// TwinCAT 3 PLC project MyLibrary
// Title: MyLibrary
// Company: FabioBolognesi
// Author: Fabio Bolognesi
// ProjectVersion: 0.0.0.0
// ProgramVersion: 3.1.4023.0
// libraries:
//   Tc2_Standard, * (Beckhoff Automation GmbH)
//   Tc2_System, * (Beckhoff Automation GmbH)
//   Tc2_Utilities, * (Beckhoff Automation GmbH)
//   Tc3_Module, * (Beckhoff Automation GmbH)
// project tree:
//   FUNCTION_BLOCKs/ FB_stringBuilder.TcPOU, FB_sweep.TcPOU, FB_timer.TcPOU
//   FUNCTIONs/ F_atan2.TcPOU, F_interpolateReal.TcPOU, F_interpolateTime.TcPOU, F_saturation.TcPOU, F_time2seconds.TcPOU, F_seconds2time.TcPOU
//   GLOBAL_VARIABLEs/ CONSTANTS.TcGVL, CONVERSIONS.TcGVL, PARAMETERs.TcGVL
//   STRUCTUREs/ ST_TypeSizes.TcDUT
// real-time tasks:
//   TASK PlcTask: cycle T#10ms, priority 20, ADS port 350

// ---- STRUCTUREs/ST_TypeSizes.TcDUT
TYPE ST_TypeSizes :
STRUCT
	// MEMORIA
	uiBIT		:	UINT	:=	SIZEOF(BIT);
	uiByte		:	UINT	:=	SIZEOF(BYTE);
	uiWord		:	UINT	:=	SIZEOF(WORD);
	uiDWord		:	UINT	:=	SIZEOF(DWORD);
	uiLWord		:	UINT	:=	SIZEOF(LWORD);
	
	// BOOL
	uiBool		:	UINT	:=	SIZEOF(BOOL);
	
	// UINTERI
	uiSUINT		:	UINT	:=	SIZEOF(SINT);
	uiUSUINT	:	UINT	:=	SIZEOF(USINT);
	uiUINT		:	UINT	:=	SIZEOF(UINT);
	uiUUINT		:	UINT	:=	SIZEOF(UINT);
	uiDUINT		:	UINT	:=	SIZEOF(DINT);
	uiUDUINT	:	UINT	:=	SIZEOF(UDINT);
	uiLUINT		:	UINT	:=	SIZEOF(LINT);
	uiULUINT	:	UINT	:=	SIZEOF(ULINT);
	
	// REALI
	uiReal		:	UINT	:=	SIZEOF(REAL);
	uiLReal		:	UINT	:=	SIZEOF(LREAL);
	
	// STRINGE
	
	// TEMPI E DATE
	uiTime		:	UINT	:=	SIZEOF(TIME);
	uiLTime		:	UINT	:=	SIZEOF(LTIME);
	uiDate		:	UINT	:=	SIZEOF(DATE);
	
	// MIE FUNCTION BLOCKS
	uiStringBuilder	:	UINT	:=	SIZEOF(FB_stringBuilder);
	uiTimer			:	UINT	:=	SIZEOF(FB_timer);
	
END_STRUCT
END_TYPE

// ---- GLOBAL_VARIABLEs/CONSTANTS.TcGVL
{attribute 'qualified_only'}
VAR_GLOBAL CONSTANT
	// ACCELERAZIONE DI GRAVITà
	G	:	REAL	:=	9.80665;
	
	// PI GRECO
	PI	:	REAL	:=	3.141592;
	
END_VAR

// ---- GLOBAL_VARIABLEs/CONVERSIONS.TcGVL
{attribute 'qualified_only'}
VAR_GLOBAL CONSTANT
	rTime2Seconds	:	REAL	:=	0.001;
	rSeconds2Time	:	REAL	:=	1000;
END_VAR

// ---- GLOBAL_VARIABLEs/PARAMETERs.TcGVL
{attribute 'global_init_slot' := '40001'}
{attribute 'qualified_only'}
VAR_GLOBAL CONSTANT
	// CARATTERI MASSIMI PER STRINGHE
	uiMaxCharacters	:	UINT	:=	5000;
END_VAR

// ---- FUNCTION_BLOCKs/FB_stringBuilder.TcPOU
FUNCTION_BLOCK FB_stringBuilder
VAR_INPUT
END_VAR
VAR
	bBuffer				:	ARRAY[0..PARAMETERS.uiMaxCharacters - 1] OF BYTE;
	bBufferOld			:	ARRAY[0..PARAMETERS.uiMaxCharacters - 1] OF BYTE;
	udiIndex			:	UDINT;
	udiIndexOld			:	UDINT;
	pbBuffer			:	POINTER TO BYTE		:=	ADR(bBuffer);
	pbBufferOld			:	POINTER TO BYTE		:=	ADR(bBufferOld);
END_VAR

METHOD AddChar : BOOL
VAR_INPUT
	byChar	:	BYTE;
END_VAR
IF CheckLength() THEN
	bBuffer[udiIndex]	:=	byChar;
	AddChar			:=	TRUE;
	IncrementIndex();
END_IF
END_METHOD

ACTION AddCloseBracket:
AddChar(41);
END_ACTION

ACTION AddColon:
AddChar(58);
END_ACTION

ACTION AddComma:
AddChar(44);
END_ACTION

ACTION AddDollar:
AddChar(36);
END_ACTION

ACTION AddDot:
AddChar(46);
END_ACTION

ACTION AddDoubleQuote:
AddChar(34);
END_ACTION

METHOD AddKeyValue : BOOL
VAR_INPUT
	psKey	:	POINTER TO STRING;
	psValue	:	POINTER TO STRING;
END_VAR
AddString(psKey);
AddColon();
AddString(psValue);
AddComma();
END_METHOD

ACTION AddNewLine:
AddChar(10);
END_ACTION

ACTION AddNullChar:
IF NOT CheckLength() THEN
	udiIndex	:=	PARAMETERS.uiMaxCharacters - 1;
END_IF
AddChar(0);
END_ACTION

ACTION AddOpenBracket:
AddChar(40);
END_ACTION

ACTION AddQuote:
AddChar(39);
END_ACTION

ACTION AddSemicolon:
AddChar(59);
END_ACTION

ACTION AddSpace:
AddChar(32);
END_ACTION

METHOD AddString : BOOL
VAR_INPUT
	psString		:	POINTER TO STRING;
END_VAR
VAR
	udiLen	:	UDINT;
END_VAR
udiLen	:=	(LEN2(psString));
IF CheckFinalLength(udiLen) THEN
	MEMCPY(pbBuffer + udiIndex, psString, udiLen);
	IncrementIndexVariable(udiLen);
	AddString	:=	TRUE;
END_IF
END_METHOD

ACTION AddTab:
AddChar(9);
END_ACTION

ACTION AddUnderscore:
AddChar(95);
END_ACTION

METHOD BuildString : BOOL
VAR_INPUT
	psString	:	POINTER TO STRING;
END_VAR
AddNullChar();
MEMCPY( psString, ADR(bBuffer), udiIndex );
END_METHOD

METHOD CheckFinalLength : BOOL
VAR_INPUT
	udiLen	:	UDINT;
END_VAR
CheckFinalLength	:=	(udiIndex + udiLen) < PARAMETERS.uiMaxCharacters;
END_METHOD

METHOD CheckLength : BOOL
VAR_INPUT
END_VAR
CheckLength	:=	CheckFinalLength(0);
END_METHOD

METHOD CheckMinimumLength : BOOL
VAR_INPUT
END_VAR
CheckMinimumLength	:=	udiIndex > 0;
END_METHOD

ACTION DecrementIndex:
IF CheckMinimumLength() THEN
	udiIndex	:=	udiIndex - 1;
END_IF
END_ACTION

METHOD DeleteChars : BOOL
VAR_INPUT
	udiNumChars	:	UDINT;
END_VAR
udiNumChars	:=	MIN(udiNumChars, udiIndex);
MEMSET(pbBuffer + (udiIndex - udiNumChars), 0, udiNumChars);
udiIndex := udiIndex - udiNumChars;
END_METHOD

ACTION IncrementIndex:
IncrementIndexVariable(1);
END_ACTION

METHOD IncrementIndexVariable : BOOL
VAR_INPUT
	udiIncrement	:	UDINT;
END_VAR
udiIndex	:=	udiIndex + udiIncrement;
END_METHOD

ACTION ResetBuffer:
IF CheckMinimumLength() THEN
	udiIndexOld	:=	udiIndex - 1;
	MEMSET(	ADR(bBufferOld), 0, PARAMETERS.uiMaxCharacters);
	MEMCPY( ADR(bBufferOld), ADR(bBuffer), udiIndexOld);
	
	ResetIndex();
	MEMSET(	ADR(bBuffer), 0, PARAMETERS.uiMaxCharacters);
END_IF
END_ACTION

ACTION ResetIndex:
udiIndex	:=	0;
END_ACTION

END_FUNCTION_BLOCK

// ---- FUNCTION_BLOCKs/FB_sweep.TcPOU
FUNCTION_BLOCK FB_sweep
VAR
	// VALORI DI INIZIALIZZAZIONE
	rStartFreq	:	REAL;
	rEndFreq	:	REAL;
	rLength		:	REAL;
	rK			:	REAL;
	
	// TIMER
	fbTimer			:	FB_Timer(T#0S);
END_VAR

METHOD ComputeFrequency : REAL
VAR_INPUT
END_VAR
ComputeFrequency	:=	F_interpolateReal(
	rX_Old	:=	0,
	rX_New	:=	rLength,
	rY_Old	:=	rStartFreq,
	rY_New	:=	rEndFreq,
	rX		:=	fbTimer.ComputeElapsedSeconds()
	);
END_METHOD

METHOD Initialize : BOOL
VAR_INPUT
	rInputStartFrequency	:	REAL;
	rInputEndFrequency		:	REAL;
	rInputLength			:	REAL;
END_VAR
rStartFreq	:=	rInputStartFrequency;
rEndFreq	:=	rInputEndFrequency;
rLength		:=	rInputLength;
rK			:=	(rEndFreq - rStartFreq) / rLength;

fbTimer.ChangeTimer(F_seconds2Time(rLength));
END_METHOD

ACTION Start:
fbTimer.Reset();
END_ACTION

METHOD Step : REAL
VAR_INPUT
END_VAR
VAR
	rTime	:	REAL;
END_VAR
IF fbTimer.VerifySelfElapsed() THEN
	Step	:=	0;
ELSE
	rTime	:=	fbTimer.ComputeElapsedSeconds();
	Step	:=	SIN(CONSTANTS.PI * rTime * (2 * rStartFreq + rK * rTime));
END_IF
END_METHOD

END_FUNCTION_BLOCK

// ---- FUNCTION_BLOCKs/FB_timer.TcPOU
FUNCTION_BLOCK FB_timer
VAR_INPUT
	tTimer		:	TIME;
END_VAR
VAR
	tStartTime	:	TIME	:=	TIME() - tTimer;
END_VAR

METHOD ChangeTimer : BOOL
VAR_INPUT
	tTimerNew	:	TIME;
END_VAR
tTimer	:=	tTimerNew;
END_METHOD

METHOD ComputeElapsed : TIME
ComputeElapsed	:=	TIME() - tStartTime;
END_METHOD

METHOD ComputeElapsedSeconds : REAL
VAR_INPUT
END_VAR
ComputeElapsedSeconds	:=	F_time2seconds(ComputeElapsed());
END_METHOD

ACTION Reset:
tStartTime	:=	TIME();
END_ACTION

METHOD ResetCondition : BOOL
VAR_INPUT
	bCondition	:	BOOL;
END_VAR
IF bCondition THEN
	Reset();
END_IF
END_METHOD

METHOD ResetWithOffset : BOOL
VAR_INPUT
	tOffset	:	TIME;
END_VAR
tStartTime	:=	TIME() - tOffset;
END_METHOD

METHOD VerifyElapsed : BOOL
VAR_INPUT
	tInputTime	:	TIME;
END_VAR
VerifyElapsed	:=	ComputeElapsed() > tInputTime;
END_METHOD

METHOD VerifySelfElapsed : BOOL
VerifySelfElapsed	:=	ComputeElapsed() > tTimer;
END_METHOD

END_FUNCTION_BLOCK

// ---- FUNCTIONs/F_time2seconds.TcPOU
FUNCTION F_time2seconds : REAL
VAR_INPUT
	tTime	:	TIME;
END_VAR
VAR
END_VAR

F_time2seconds	:=	TIME_TO_REAL(tTime) * CONVERSIONS.rTime2Seconds;

END_FUNCTION

// ---- FUNCTIONs/F_interpolateReal.TcPOU
FUNCTION F_interpolateReal : REAL
VAR_INPUT
	rX_Old	:	REAL;
	rX_New	:	REAL;
	rY_Old	:	REAL;
	rY_New	:	REAL;
	rX		:	REAL;
END_VAR
VAR
END_VAR

IF rX_Old <> rX_New THEN
	IF rX < rX_Old THEN
		F_interpolateReal	:=	rY_Old;
	ELSIF rX > rX_New THEN
		F_interpolateReal	:=	rY_New;
	ELSE
		F_interpolateReal	:=	rY_Old + (rY_New - rY_Old) / (rX_New - rX_Old) * (rX - rX_Old);
	END_IF
ELSE
	F_interpolateReal	:=	0;
END_IF

END_FUNCTION

// ---- FUNCTIONs/F_seconds2time.TcPOU
FUNCTION F_seconds2time : TIME
VAR_INPUT
	rSeconds	:	REAL;
END_VAR
VAR
END_VAR

F_seconds2time	:=	REAL_TO_TIME(rSeconds * CONVERSIONS.rSeconds2Time);

END_FUNCTION

// ---- FUNCTIONs/F_atan2.TcPOU
FUNCTION F_atan2 : REAL
VAR_INPUT
	rX	:	REAL;
	rY	:	REAL;
END_VAR
VAR
END_VAR

// CALCOLO L'ANGOLO CONOSCENDO COORDINATE X E Y
IF rX > 0 THEN
	F_atan2	:=	ATAN(rY / rX);
ELSIF rX = 0 AND rY > 0 THEN
	F_atan2	:=	LREAL_TO_REAL(CONSTANTS.PI / 2);
ELSIF rX = 0 AND rY < 0 THEN
	F_atan2	:=	- LREAL_TO_REAL(CONSTANTS.PI / 2);
ELSIF rX < 0 AND rY >= 0 THEN
	F_atan2	:=	LREAL_TO_REAL(ATAN(rY / rX) + CONSTANTS.PI);
ELSIF rX < 0 AND rY < 0 THEN
	F_atan2	:=	LREAL_TO_REAL(ATAN(rY / rX) - CONSTANTS.PI);
END_IF

END_FUNCTION

// ---- FUNCTIONs/F_interpolateTime.TcPOU
FUNCTION F_interpolateTime : REAL
VAR_INPUT
	tX_Old	:	TIME;
	tX_New	:	TIME;
	rY_Old	:	REAL;
	rY_New	:	REAL;
	tX		:	TIME;
END_VAR
VAR
END_VAR

F_interpolateTime	:=	F_interpolateReal(
	rX_Old	:=	F_time2seconds(tX_Old),
	rX_New	:=	F_time2seconds(tX_New),
	rY_Old	:=	rY_Old,
	rY_New	:=	rY_New,
	rX		:=	F_time2seconds(tX)
	);

END_FUNCTION

// ---- FUNCTIONs/F_saturation.TcPOU
FUNCTION F_saturation : REAL
VAR_INPUT
	rInput			:	REAL;
	rMinimumValue	:	REAL;
	rMaximumValue	:	REAL;
END_VAR
VAR
END_VAR

// ESEGUO UNA SATURAZIONE DEL VALORE IN INGRESSO
F_saturation	:=	MAX(rMinimumValue, MIN(rMaximumValue, rInput));

END_FUNCTION
